FUNCTION_BLOCK FB_Conveyor
VAR
    motor : I_Motor;
    requested : BOOL;
    configuredDelay : TIME := T#100ms;
    speed : LREAL := 0.5;
    count : UDINT;
    alarmText : STRING(80);
END_VAR

(* Methods control the dependency explicitly. *)

METHOD PUBLIC BindMotor
VAR_INPUT
    motor : I_Motor;
END_VAR
(* Stop the old dependency before replacing it; a new Start is required. *)
IF THIS^.motor <> 0 THEN
    THIS^.motor.Update(run := FALSE, delay := configuredDelay);
END_IF;
THIS^.motor := motor;
requested := FALSE;
END_METHOD

METHOD PUBLIC Start
VAR_INPUT
    delay : TIME := T#100ms;
END_VAR
configuredDelay := delay;
requested := TRUE;
END_METHOD

METHOD PUBLIC Stop
requested := FALSE;
IF motor <> 0 THEN
    motor.Update(run := FALSE, delay := configuredDelay);
END_IF;
alarmText := 'Stopped';
END_METHOD

METHOD PUBLIC Update
VAR_INPUT
    guardClosed : BOOL;
    stopRequested : BOOL := FALSE;
    sensor : BOOL := FALSE;
END_VAR
VAR_INST
    productEdge : R_TRIG;
END_VAR
productEdge(CLK := sensor);
IF motor = 0 THEN
    requested := FALSE;
    alarmText := 'Motor not bound';
    RETURN;
END_IF;
IF stopRequested OR NOT guardClosed OR motor.Faulted THEN
    requested := FALSE;
END_IF;
motor.SpeedSetpoint := speed;
motor.Update(run := requested, delay := configuredDelay);
IF motor.Running AND productEdge.Q THEN
    count := count + 1;
END_IF;
IF NOT guardClosed THEN
    alarmText := 'Guard open';
ELSIF stopRequested THEN
    alarmText := 'Stopped';
ELSIF motor.Faulted THEN
    alarmText := 'Motor fault';
ELSIF requested AND NOT motor.Running THEN
    alarmText := 'Starting';
ELSE
    alarmText := '';
END_IF;
END_METHOD

PROPERTY PUBLIC SpeedSetpoint : LREAL
GET
SpeedSetpoint := THIS^.speed;
END_GET
SET
THIS^.speed := LIMIT(0.0, SpeedSetpoint, 1.0);
END_SET
END_PROPERTY

PROPERTY PUBLIC Running : BOOL
GET
IF motor <> 0 THEN
    Running := motor.Running;
END_IF;
END_GET
END_PROPERTY

PROPERTY PUBLIC ActiveSpeed : LREAL
GET
IF motor <> 0 THEN
    ActiveSpeed := motor.ActualSpeed;
END_IF;
END_GET
END_PROPERTY

PROPERTY PUBLIC ProductCount : UDINT
GET
ProductCount := count;
END_GET
END_PROPERTY

PROPERTY PUBLIC Alarm : STRING(80)
GET
Alarm := alarmText;
END_GET
END_PROPERTY

END_FUNCTION_BLOCK

(* stored: Version 1.1.0.1, ProductVersion 3.1 *)
